INTERFACE I_Alarm

METHOD addAlarm : BOOL
VAR_INPUT
	sKoodi		: STRING;
	sKuvaus		: STRING;
END_VAR
END_METHOD

END_INTERFACE

(* stored: Version 1.1.0.1
   Itf I_Alarm: Id {70f374ee-1dca-4b66-b1b4-e7b455663b12}
   Method addAlarm: Id {39386a93-8060-4c8c-926d-f614b9016e67} *)
